INTERFACE I_Valve

METHOD Open : BOOL
END_METHOD

PROPERTY State : E_ValveState
GET
END_GET
SET
END_SET
END_PROPERTY

END_INTERFACE

(* stored: Version 1.1.0.1, ProductVersion 3.1.4024.12
   Itf I_Valve: Id {fbaa47fe-d0d9-42e9-91ce-6670802fec89}
   Method Open: Id {5328a085-5906-42d7-8998-6e575ad59e3c}
   Property State: Id {f73f887f-087b-4edc-b5b2-8ce8f0dfad06}
   Get Get: Id {8f7ea9e1-0a9d-41ac-b57b-61ed5fc58b3b}
   Set Set: Id {6d6ce055-980f-4bee-aab4-a282cee0e164} *)
